(* IEC 61131-3 sources: codesys-framework/txt/application/WeVe Core (library)/60 Event/I_EventGroup, 5 files *)

(* ---- Condition.method.st ---- *)
// Doorgeefluik naar I_Event.Condition van event iEvent (enum van de eigenaar).
// Geeft Active van dat event terug, FALSE bij een ongeldige index.
METHOD Condition : BOOL
VAR_INPUT
	iEvent 			: INT;
	xCondition 		: BOOL;
	scPayload 		: SC_EventPayload := (asPayload := [10('')]);	// mag weggelaten worden
END_VAR

(* ---- GetEvent.method.st ---- *)
// Rechtstreekse toegang tot één event, voor uitzonderlijke gevallen.
// Geeft 0 terug bij een ongeldige index: altijd controleren op <> 0.
METHOD GetEvent : I_Event
VAR_INPUT
	iEvent 			: INT;
END_VAR

(* ---- Initialize.method.st ---- *)
// Config van alle events invullen en de logger doorgeven. Eenmalig, in de eerste cyclus.
// TRUE = klaar.
METHOD Initialize : BOOL
VAR_INPUT
END_VAR

(* ---- Log.method.st ---- *)
// Doorgeefluik naar I_Event.Log van event iEvent (enum van de eigenaar).
// FALSE bij een ongeldige index.
METHOD Log : BOOL
VAR_INPUT
	iEvent 			: INT;
	scPayload 		: SC_EventPayload := (asPayload := [10('')]);	// mag weggelaten worden
END_VAR

(* ---- Reset.method.st ---- *)
// Reset alle events van de groep. TRUE = geen enkel event nog actief.
METHOD Reset : BOOL
VAR_INPUT
END_VAR
